TYPE ST_Array :
STRUCT
	arr1 : ARRAY[0..2,0..2] OF INT;
	arr2 : ARRAY[0..1,0..1] OF ARRAY[0..1,0..1] OF INT;
	arr3 : ARRAY[0..1,0..1,0..1] OF ARRAY[0..1] OF INT;
END_STRUCT
END_TYPE

(* stored: Version 1.1.0.1, ProductVersion 3.1.4026.19
   DUT ST_Array: Id {c5e05f51-855c-4d14-af57-4b9f77fa44de} *)
